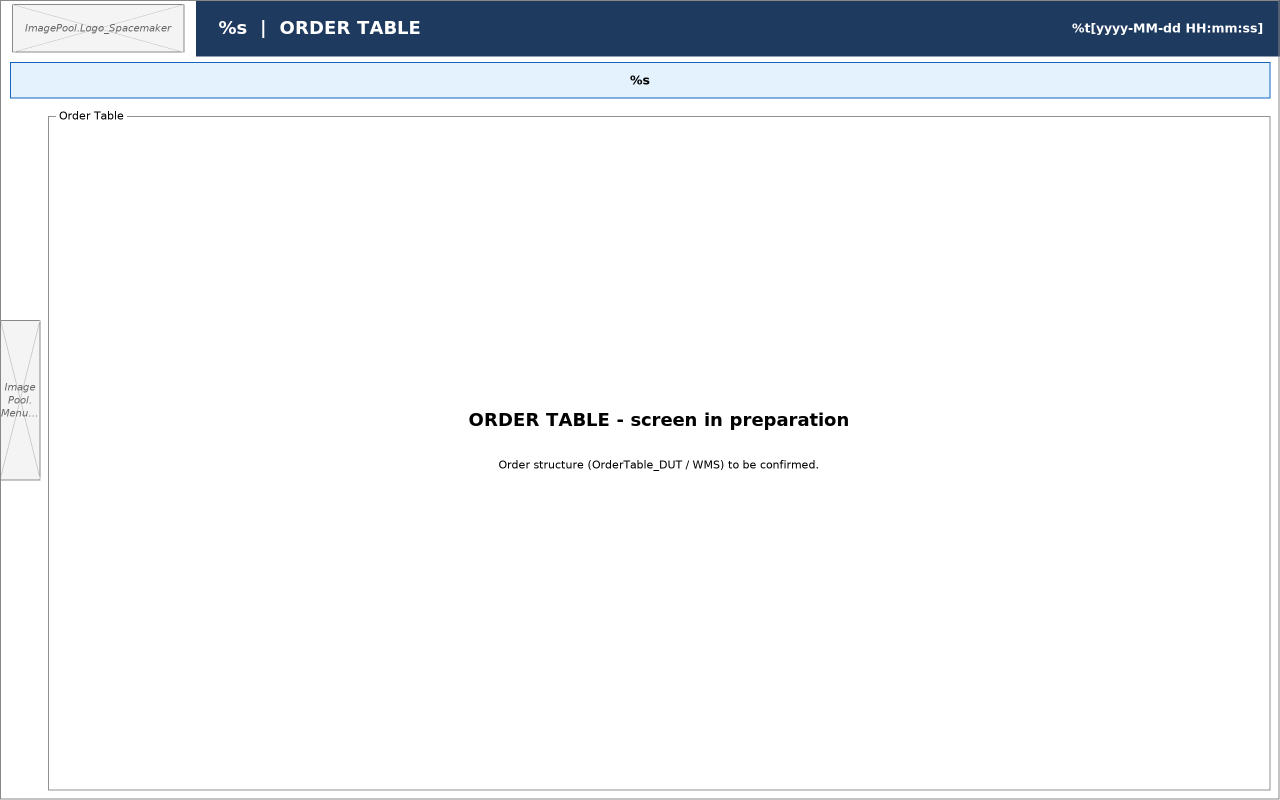
VISUALIZATION Order_Table  // 1280x800
    Rectangle (0,0 196x56)
        OnMouseClick: change screen: Main
    Image (12,4 172x48), image: ImagePool.Logo_Spacemaker
        OnMouseClick: change screen: Main
    Rectangle (196,0 1084x56), "%s | ORDER TABLE", text variable: GVL_HMI_System.stStatus.sSystemName
    Rectangle (930,8 336x40), "%t[yyyy-MM-dd HH:mm:ss]", text variable: GVL_HMI_System.stStatus.dtNow
    Rectangle (10,62 1260x36), "%s", text variable: GVL_HMI_System.stStatus.sMessage, colour toggle: GVL_HMI_System.stStatus.bMessageAlarm
    GroupBox (48,108 1222x682), "Order Table"
    Rectangle (78,400 1162x40), "ORDER TABLE - screen in preparation"
    Rectangle (78,450 1162x30), "Order structure (OrderTable_DUT / WMS) to be confirmed."
    Rectangle (0,320 40x160)
        OnMouseEnter: OpenDialog Dialog=Dialog, OpenModal=True, PositionX=0, PositionY=0
        OnMouseClick: OpenDialog Dialog=Dialog, OpenModal=True, PositionX=0, PositionY=0
    Image (0,320 40x160), image: ImagePool.Menu_Tab
        OnMouseEnter: OpenDialog Dialog=Dialog, OpenModal=True, PositionX=0, PositionY=0
        OnMouseClick: OpenDialog Dialog=Dialog, OpenModal=True, PositionX=0, PositionY=0
END_VISUALIZATION

(* stored: Version 1.1.0.1
   Visu Order_Table: Id {12c7abed-f61d-4ccb-95bd-df0ffe4e3346} *)
